// TIA Portal V19 export
DATA_BLOCK "AI_TT02"   // DB5
// stored: InstanceOfName AI, InstanceOfType FB
"AI"
   // VAR_INPUT
   //    RAW_MIN : Int;
   //    RAW_MAX : Int;
   //    SCALE_MIN : Real;
   //    SCALE_MAX : Real;
   //    HH_SP : Real;
   //    HSP : Real;
   //    LL_SP : Real;
   //    LSP : Real;
   //    ALM_WT : Time;
   //    INPUT : Int;
   // END_VAR
   // VAR_OUTPUT
   //    FAULT : Bool;
   //    HH_ALM : Bool;
   //    H_ALM : Bool;
   //    LL_ALM : Bool;
   //    L_ALM : Bool;
   //    SCALE_OUT : Real;
   // END_VAR
   // VAR
   //    AI : "SCALING";
   //    MAX_VALUE : Int;
   //    HH_TIME { S7_SetPoint := 'True'} : TON_TIME;
   //    H_TIME { S7_SetPoint := 'True'} : TON_TIME;
   //    LL_TIME { S7_SetPoint := 'True'} : TON_TIME;
   //    L_TIME { S7_SetPoint := 'True'} : TON_TIME;
   // END_VAR
BEGIN
END_DATA_BLOCK
